Yaskawa INFORM job: SPEEDPR.JBI

/JOB
//NAME SPEEDPR
//POS
///NPOS 21,0,21,0,0,0
///TOOL 9
///POSTYPE PULSE
///PULSE
C00000=0,0,0
C00001=0,0,0
C00002=0,0,0
C00003=0,0,0
C00004=0,0,0
C00005=0,0,0
C00006=0,0,0
C00007=0,0,0
C00008=0,0,0
C00009=0,0,0
C00010=0,0,0
C00011=0,0,0
C00012=0,0,0
C00013=0,0,0
C00014=0,0,0
C00015=0,0,0
C00016=0,0,0
C00017=0,0,0
C00018=0,0,0
C00019=0,0,0
C00020=0,0,0
EC00000=0
EC00001=0
EC00002=0
EC00003=0
EC00004=0
EC00005=0
EC00006=0
EC00007=0
EC00008=0
EC00009=0
EC00010=0
EC00011=0
EC00012=0
EC00013=0
EC00014=0
EC00015=0
EC00016=0
EC00017=0
EC00018=0
EC00019=0
EC00020=0
//INST
<volatile>
///COMM Generated using RoboDK
///ATTR SC,RW
///GROUP1 RB1
NOP
'Program generated by RoboDK v
'6.0.7 for Yaskawa Motoman EPL
'160 on XX/XX/XXXX 18:00:00
'Using nominal kinematics.
'Using Frame S (targets wrt ba
'se):
'1234.6,-98.8,50.5,0.0,0.0,30.
'0
'Tool Tool S should be close t
'o:
'10.0,20.0,150.0,0.0,0.0,0.0
MOVL C00000 V=1.0 PL=0  +MOVJ EC00000 VJ=100.00
MOVJ C00001 VJ=1.00 PL=0  +MOVJ EC00001 VJ=100.00
MOVL C00002 V=12.3 PL=1  +MOVJ EC00002 VJ=100.00
MOVJ C00003 VJ=5.50 PL=1  +MOVJ EC00003 VJ=100.00
MOVL C00004 V=99.9 PL=2  +MOVJ EC00004 VJ=100.00
MOVJ C00005 VJ=20.00 PL=2  +MOVJ EC00005 VJ=100.00
MOVL C00006 V=333.3 PL=4  +MOVJ EC00006 VJ=100.00
MOVJ C00007 VJ=45.00 PL=4  +MOVJ EC00007 VJ=100.00
MOVL C00008 V=1000.0 PL=6  +MOVJ EC00008 VJ=100.00
MOVJ C00009 VJ=90.00 PL=6  +MOVJ EC00009 VJ=100.00
MOVL C00010 V=2000.0 PL=8  +MOVJ EC00010 VJ=100.00
MOVJ C00011 VJ=100.0 PL=8  +MOVJ EC00011 VJ=100.00
MOVL C00012 V=2000.0 PL=8  +MOVJ EC00012 VJ=100.00
MOVJ C00013 VJ=100.0 PL=8  +MOVJ EC00013 VJ=100.00
MOVL C00014 V=2000.0 PL=8  +MOVJ EC00014 VJ=100.00
MOVJ C00015 VJ=100.0 PL=8  +MOVJ EC00015 VJ=100.00
MOVL C00016 V=0.5 PL=8  +MOVJ EC00016 VJ=100.00
MOVJ C00017 VJ=100.0 PL=8  +MOVJ EC00017 VJ=100.00
MOVL C00018 V=750.0 PL=8  +MOVJ EC00018 VJ=100.00
MOVJ C00019 VJ=2.25 PL=8  +MOVJ EC00019 VJ=100.00
MOVL C00020 V=750.0  +MOVJ EC00020 VJ=100.00
END
